(* IEC 61131-3 sources: JingjiangMoonbox/Application/Application/任务列表/OtherTask, 5 files *)

(* ---- KS_ArcFollow1UFlag_Deal.st ---- *)
(*@CES
Name=KS_ArcFollow1UFlag_Deal
Type=FunctionBlock
TypeGuid=6f9dac99-8de1-4efc-8465-68ac443b7d08
Guid=d7f43731-9672-42b8-a130-8c9a3b5ea44f
HasDeclaration=True
HasImplementation=True
*)
{DECLARATION}
FUNCTION KS_ArcFollow1UFlag_Deal : BOOL(*所有套色跟踪第一色标志处理@优化为了跟踪任意色@2024.02.22.102708*)
(*输出的标志可能决定了是否打开双波门*)
(*套色误差到达一定阈值时输出跟踪第一色标志-置位后就不再复位除非关闭使能
@用于解决在拉伸比较大的材料上后面色组找不到1色的问题。
@最大16个轴@c_byAxisNum_Max 确定*)
(*2024.02.22.085437 将检查第一个套色轴修改为检查跟踪的套色轴的下一个轴的误差*)
(*2025.1.9.145517 增加套色轴到达误差范围标志*)
VAR_INPUT
	i_xEn:BOOL;(*处理使能*)
	i_byArcNum_Max:BYTE;(*最大套色轴个数@最大16个*)
	i_byGrpAxisNum_Pu:BYTE;(*系中色组轴个数*)
	i_pabyGrpAxisList:POINTER TO BYTE;(*系的轴ID列表首地址*)
	i_byArcNum:BYTE;(*当前套色轴个数*)
	i_pabyArcAxisList:POINTER TO BYTE;(*套色的轴列表首地址@2024.02.22.084654*)
	i_pabyArcIdList:POINTER TO BYTE;(*套色的ID列表首地址*)
	i_byArcErr_Threshold:BYTE:=50;(*套色误差阈值@单位丝*)
	i_byContinuousCycleCnt:BYTE:=10;(*持续的圈数@持续这么多幅误差都在阈值以内就认为可以输出标志*)
	i_paxArcErrValid:POINTER TO ARRAY [1..c_byAxisNum_Max] OF BOOL;(*误差值有效了*)
	i_aiArcErr:ARRAY [1..c_byAxisNum_Max] OF INT;(*套色误差值(在让料头未到达的时候误差值写成最大值)@索引为色组号*)
	i_pabyCycleCnt:POINTER TO ARRAY [1..c_byAxisNum_Max] OF BYTE;(*满足条件后的圈数计数值@索引为色组号*)
	i_paxArcReachRangeFlag:POINTER TO ARRAY [1..c_byAxisNum_Max] OF BOOL;(*套色到达阈值标志@用于判断是否要输出跟踪第一色标志*)
	i_paxArcFollow1UFlag:POINTER TO ARRAY [1..c_byAxisNum_Max] OF BOOL;(*输出跟踪第一色标志@索引为色组号*)
	i_pabyFollowArcId:POINTER TO ARRAY [1..c_byAxisNum_Max] OF BYTE;(*2024.02.22.100117 跟踪的套色id@索引为轴id*)
	i_pxArcErrInRange:POINTER TO BOOL;(*套色误差在范围内@2025.1.9.145628+*)
END_VAR
VAR
	iN: INT;
	iM: INT;
	iAxisId: INT;
	iArcId: INT;
	byArcNum_Max: BYTE;
	byArcErr_Threshold: BYTE;(*丝单位*)
	byContinuousCycleCnt: BYTE;(*持续的幅数计数值*)

	byGrpAxisNum_Pu: BYTE;
	pabyGrpAxisList_Tmp:POINTER TO ARRAY [1..c_byAxisNum_Max] OF BYTE;(*系轴id列表*)
	abyGrpAxisList:ARRAY [1..c_byAxisNum_Max] OF BYTE;(*系轴id列表*)

	byArcNum: BYTE;
	pabyArcAxisList_Tmp:POINTER TO ARRAY [1..c_byAxisNum_Max] OF BYTE;(*套色轴id列表*)
	abyArcAxisList:ARRAY [1..c_byAxisNum_Max] OF BYTE;(*套色轴id列表*)
	pabyArcIdList_Tmp:POINTER TO ARRAY [1..c_byAxisNum_Max] OF BYTE;(*套色轴色序id列表*)
	abyArcIdList:ARRAY [1..c_byAxisNum_Max] OF BYTE;(*套色轴色序id列表*)
	axArcReachRangeFlag:ARRAY [1..c_byAxisNum_Max] OF BOOL;(*套色到达阈值标志*)
	axArcFollow1UFlag:ARRAY [1..c_byAxisNum_Max] OF BOOL;(*输出跟踪第一色标志@索引为色组号*)
	abyCycleCnt:ARRAY [1..c_byAxisNum_Max] OF BYTE;(*每个轴的循环计数*)
	aiArcErr:ARRAY [1..c_byAxisNum_Max] OF INT;(*套色误差*)
	axNeedRstAxisId: ARRAY [1..c_byAxisNum_Max] OF BOOL;(*需要复位参数的轴id|默认写true'*)
	axArcErrValid: ARRAY [1..c_byAxisNum_Max] OF BOOL;(*套色误差有效标志位*)
	xArvErrValid: BOOL;(*误差都有效了-可以检查标志*)
	xFollow1UEn: BOOL;(*跟踪第一色使能了*)

	abyFollowArcId:ARRAY [1..c_byAxisNum_Max] OF BYTE;(*2024.02.22.100 跟踪的套色id*)
	iFollowArcId:INT;
	iCheckArcIdSa:INT;(*开始检查的套色id*)
	iIndex: INT;
	iArcErrInRangeAxisCnt: INT;(*在范围的轴个数@2025.1.9.145758*)
END_VAR

VAR CONSTANT
	(*修改的时候谨慎点@外面输入的都是16个轴*)
	c_byAxisNum_Max:BYTE:=16;(*最大的轴个数@直接写死*)
END_VAR
{IMPLEMENTATION}
byArcNum_Max:=i_byArcNum_Max;
IF byArcNum_Max=0 OR
	byArcNum_Max>c_byAxisNum_Max THEN
	byArcNum_Max:=c_byAxisNum_Max;
END_IF

byArcNum:=i_byArcNum;
IF byArcNum>c_byAxisNum_Max THEN
	byArcNum:=c_byAxisNum_Max;
END_IF

byGrpAxisNum_Pu:=i_byGrpAxisNum_Pu;
IF byGrpAxisNum_Pu>c_byAxisNum_Max THEN
	byGrpAxisNum_Pu:=c_byAxisNum_Max;
END_IF

byArcErr_Threshold:=i_byArcErr_Threshold;
byContinuousCycleCnt:=i_byContinuousCycleCnt;

IF i_paxArcErrValid<>0 THEN
	axArcErrValid:=i_paxArcErrValid^;
END_IF
aiArcErr:=i_aiArcErr;

(*获取系轴列表信息*)
IF i_pabyGrpAxisList<>0 THEN
	pabyGrpAxisList_Tmp:=i_pabyGrpAxisList;
	abyGrpAxisList:=pabyGrpAxisList_Tmp^;
END_IF

(*获取套色轴列表信息*)
IF i_pabyArcAxisList<>0 THEN
	pabyArcAxisList_Tmp:=i_pabyArcAxisList;
	abyArcAxisList:=pabyArcAxisList_Tmp^;
END_IF

IF i_pabyArcIdList<>0 THEN
	pabyArcIdList_Tmp:=i_pabyArcIdList;
	abyArcIdList:=pabyArcIdList_Tmp^;
END_IF

IF i_pabyCycleCnt<>0 THEN
	abyCycleCnt:=i_pabyCycleCnt^;
END_IF
IF i_paxArcReachRangeFlag <>0 THEN
	axArcReachRangeFlag:=i_paxArcReachRangeFlag^;
END_IF
IF i_paxArcFollow1UFlag<>0 THEN
	axArcFollow1UFlag:=i_paxArcFollow1UFlag^;
END_IF

IF i_pabyFollowArcId<>0 THEN
	abyFollowArcId:=i_pabyFollowArcId^;
END_IF

(*只处理当前系的轴*)
FOR iN:=1 TO c_byAxisNum_Max BY 1 DO(*iN为系id索引*)
	iAxisId:=abyGrpAxisList[iN];
	IF iAxisId>0 AND iAxisId<c_byAxisNum_Max THEN
		axNeedRstAxisId[iAxisId]:=TRUE;
	ELSE;(*不在这个系的轴就不管了*)
	END_IF
END_FOR

iArcErrInRangeAxisCnt:=0;
FOR iN:=2 TO byArcNum BY 1 DO(*iN为索引@从第二个套色轴开始*)
	iAxisId:=abyArcAxisList[iN];(*套色的轴id*)
	iArcId:=abyArcIdList[iN];(*套色的色序id*)
	iFollowArcId:=abyFollowArcId[iN];(*跟踪的套色Id@2024.02.22.100304*)

	IF iAxisId>=2 AND iAxisId<=c_byAxisNum_Max AND(*轴号合法@从2号轴开始*)
		iArcId>=2 AND iArcId<=c_byAxisNum_Max THEN(*色序id合法*)
		xArvErrValid:=axArcErrValid[iAxisId];(*获取误差是否有效标志位*)
		axArcErrValid[iAxisId]:=FALSE;(*使用完了就复位*)
		(*检查各个色组是否到达阈值*)
		KS_ArcAxisReachRange(
			i_xEn (*i_xEn*),
			INT_TO_BYTE(iArcId)(*i_byArcId*),
			byArcErr_Threshold(*i_byArcErr_Threshold*),
			byContinuousCycleCnt(*i_byContinuousCycleCnt*),
			xArvErrValid(*i_xArcErrValid*),
			aiArcErr[iAxisId](*i_iArcErr*),
			ADR(abyCycleCnt[iAxisId])(*i_pbyCycleCnt*),
			ADR(axArcReachRangeFlag[iAxisId])(*i_xArcReachRangeFlag*));

		(*2025.1.9.145715+*)
		IF axArcReachRangeFlag[iAxisId] THEN
			iArcErrInRangeAxisCnt:=iArcErrInRangeAxisCnt+1;
		END_IF

		(*当前色已经到达阈值了@检查之前的套色轴是否到达。确定是否要输出跟踪第一色标志*)
		IF iFollowArcId<>0 THEN(*跟踪任意色@色序id*)
			IF iArcId>2 THEN(*色序超过3的才检查别的色*)
				IF axArcReachRangeFlag[iAxisId] THEN
					(*找到跟踪的套色id在套色id列表的索引值@2024.02.22.101030+*)
					iIndex:=iN;(*非法处理@未找到色序下面判断的循环就直接跳出*)
					FOR iM:=1 TO iN-1 BY 1 DO
						IF iFollowArcId = abyArcIdList[iM]THEN
							iIndex:=iM;
							EXIT;
						END_IF
					END_FOR

					(*如果找不到,会进入下面的else分支,但是iIndex=iN|所以也不会进入循环-也就是标志不会被置位*)
					iCheckArcIdSa:=2;
					IF iIndex<>In THEN(*找到了*)
						iIndex:=iIndex+1;(*从跟踪的下一个开始检查@索引值为开始检索的值*)
						iCheckArcIdSa:=abyArcIdList[iIndex];
					END_IF

					IF iCheckArcIdSa>=iArcId THEN(*检查的值和当前的色序一样@就直接输出标志*)
						axArcFollow1UFlag[iAxisId]:=TRUE;
					ELSE(*需要经过下面的检查输出*)
						(*修改为了跟踪色+1开始@2024.02.22.104458*)
						FOR iM:=iIndex TO iN-1  BY 1 DO(*从2色色序开始检查-自己在外围条件已经检查了@im也是色序*)
							IF axArcReachRangeFlag[abyArcAxisList[iM]] THEN(*到达阈值范围了*)
								IF iM=iN-1 THEN(*前一个也到达了则输出跟踪第一色标志*)
									axArcFollow1UFlag[iAxisId]:=TRUE;
								END_IF
							ELSE(*未到达则退出循环*)
								EXIT;
							END_IF
						END_FOR
					END_IF
				ELSE
					axArcFollow1UFlag[iAxisId]:=FALSE;
				END_IF
			ELSE
				axArcFollow1UFlag[iAxisId]:=axArcReachRangeFlag[iAxisId];(*只关心自己*)
			END_IF
		ELSE(*不跟踪任意色*)
			axArcFollow1UFlag[iAxisId]:=FALSE;
		END_IF
		(*处理未套色轴-复位标志@套色轴辅助变量已经在上面清除处理了*)
		axNeedRstAxisId[iAxisId]:=FALSE;
	ELSE;(*不做处理*)
	END_IF
END_FOR
(*检查所有轴是不是都在范围内@2025.1.9.145846*)
IF i_pxArcErrInRange<>0 THEN
	IF	(iArcErrInRangeAxisCnt+1) = byArcNum AND byArcNum>1 THEN
		i_pxArcErrInRange^:=TRUE;
	ELSE
		i_pxArcErrInRange^:=FALSE;
	END_IF
END_IF

(*没处理的轴数据清除*)
FOR iAxisId:=1 TO c_byAxisNum_Max BY 1 DO
	IF axNeedRstAxisId[iAxisId] THEN
		abyCycleCnt[iAxisId]:=0;
		axArcReachRangeFlag[iAxisId]:=FALSE;
		axArcFollow1UFlag[iAxisId]:=FALSE;
		axArcErrValid[iAxisId]:=FALSE;
	END_IF
END_FOR

IF i_pabyCycleCnt<>0 THEN
	i_pabyCycleCnt^:=abyCycleCnt;
END_IF
IF i_paxArcReachRangeFlag <>0 THEN
	i_paxArcReachRangeFlag^:=axArcReachRangeFlag;
END_IF
IF i_paxArcFollow1UFlag<>0 THEN
	i_paxArcFollow1UFlag^:=axArcFollow1UFlag;
END_IF

IF i_paxArcErrValid<>0 THEN
	i_paxArcErrValid^:=axArcErrValid;
END_IF

(* ---- KS_CalcGatePos_Follow.st ---- *)
(*@CES
Name=KS_CalcGatePos_Follow
Type=FunctionBlock
TypeGuid=6f9dac99-8de1-4efc-8465-68ac443b7d08
Guid=4fe415d3-d686-4f37-995a-ecb110eaba4a
HasDeclaration=True
HasImplementation=True
*)
{DECLARATION}
FUNCTION KS_CalcGatePos_Follow : INT(*计算跟踪某一个色方式计算该色的波门位置@单位是粗采样点数*)
(*-1 参数错误
-2 标记非法
-3 未隔色*)
(*2024.02.21.130156 输出第二波们的位置@出错则输出=0*)
(*2024.7.30.144846 计算方法有问题取巧未使用实际距离使用了波门宽度@波门宽度变化为非20后就会出错了
处理为根据实际距离计算*)
(*2024.7.31.075422 2色按照波门宽度偏移*)
VAR_INPUT
	i_byUnitId_Follow:BYTE;(*跟踪的色组id*)
	i_byUnitId_Cur:BYTE;(*当前的色组id*)
	i_iGateSa:INT;(*当前波门位置*)
	i_iGateWidthRondPt:INT;(*波门宽度的粗采样点数@使用改变量需要波门宽度为20mm*)
	i_iGatePoint_Max:INT;(*最大粗采样点数*)
	i_iMarkArrangeId:INT;(*标记类型*)

	i_rGirth:REAL;(*版辊周长@mm*)
END_VAR
VAR
	byDeltaId: BYTE;
	iGateSaEx: INT;
	iRtn: INT;
	iDeltaRondPt: INT;(*间隔的粗采样点数*)
END_VAR
{IMPLEMENTATION}
IF i_iGatePoint_Max=0 THEN
	i_iGatePoint_Max:=4000;
END_IF
IF i_byUnitId_Follow>0 AND
	i_byUnitId_Cur>=2 AND(*条件修改*)
	i_byUnitId_Follow<i_byUnitId_Cur AND
	i_iGateSa>=0 AND i_iGateSa<i_iGatePoint_Max THEN

	IF i_byUnitId_Cur>i_byUnitId_Follow THEN
		byDeltaId:=i_byUnitId_Cur-i_byUnitId_Follow;(*间隔*)
	ELSE
		byDeltaId:=0;
	END_IF

	IF byDeltaId<>0 THEN;
	ELSE(*不隔色*)
		iGateSaEx:= 0;
		iRtn:=-3;
		RETURN;
	END_IF

	IF i_rGirth<>0 THEN;
	ELSE
		i_rGirth:=500;
	END_IF
	IF i_byUnitId_Cur=2 THEN(*2色按照波门宽度偏移@2024.7.31.075310*)
		iDeltaRondPt:=i_iGateWidthRondPt;
	ELSE
		iDeltaRondPt:=REAL_TO_INT(BYTE_TO_REAL(byDeltaId)*20.0/i_rGirth*i_iGatePoint_Max)+1;(*按照间隔n*20mm计算|稍微离远点@主要是1 2色的波门*)
	END_IF

	IF i_iMarkArrangeId= MARK_ARRANGE_VFOR THEN(*顺序*)
		iGateSaEx:=i_iGateSa-(*byDeltaId*i_iGateWidthRondPt*)iDeltaRondPt;
		IF iGateSaEx<0 THEN
			iGateSaEx:= iGateSaEx+i_iGatePoint_Max;
		END_IF
	ELSIF i_iMarkArrangeId= MARK_ARRANGE_VREV THEN(*逆序*)
		iGateSaEx:=i_iGateSa+(*byDeltaId*i_iGateWidthRondPt*)iDeltaRondPt;
		IF iGateSaEx>i_iGatePoint_Max THEN
			iGateSaEx:= iGateSaEx-i_iGatePoint_Max;
		END_IF
	ELSE
		iGateSaEx:= 0;
		iRtn:=-2;
	END_IF
ELSE
	iGateSaEx:= 0;
	iRtn:=-1;
END_IF
(*
IF iRtn<0 THEN
	KS_CalcGatePos_Follow:=iRtn;
ELSE*)
	KS_CalcGatePos_Follow:=iGateSaEx;
(*END_IF*)

(* ---- KS_FB_GetLatchValue.st ---- *)
(*@CES
Name=KS_FB_GetLatchValue
Type=FunctionBlock
TypeGuid=6f9dac99-8de1-4efc-8465-68ac443b7d08
Guid=ed2f2b11-af18-4922-a052-26b8330b7fb0
HasDeclaration=True
HasImplementation=True
*)
{DECLARATION}
FUNCTION_BLOCK KS_FB_GetLatchValue
VAR_INPUT
	i_xEn : BOOL;
	i_iGrpUnitNum: INT;
	i_pstStSysParam: POINTER TO StSysParam;
	i_pastStLatch : POINTER TO ARRAY [1..MAX_UNIT_NUM] OF StLatch;
END_VAR
VAR_OUTPUT
END_VAR
VAR
	iN : INT;
	iM : INT;
	iRtn : INT;
	audiTempData : ARRAY [1..MAX_UNIT_NUM] OF UDINT;
END_VAR

{IMPLEMENTATION}

IF i_xEn THEN
	IF i_pstStSysParam <> 0 AND i_pastStLatch <> 0 THEN
		FOR iN := 1 TO i_iGrpUnitNum BY 1 DO
			iRtn := GTN_GetMailbox(
				core:= 1,
				station:= 0,
				byteAddress:= 16#C412, //锁存时间32位数据（低24位锁存时间，高8位di触发次数），单位us,:低16位网络地址0xc412,高16位网络地址0xc414
				pData:= ADR(audiTempData[iN]),
				wordCount:= 2,
				dataMode:= 1,
				desId:=iN,
				typeVar:= 1);

			i_pastStLatch^[iN].iTriggerCnt := UDINT_TO_INT(SHR(audiTempData[iN],24));
			i_pastStLatch^[iN].udiTriggerTimeErr := SHR(SHL(audiTempData[iN],16#8),16#8);

			iRtn := GTN_GetMailbox(
				core:= 1,
				station:= 0,
				byteAddress:= 16#C454, //锁存编码器32位数据，一个版周最大脉冲值131072，低16位网络地址0xc454，高16位网络地址0xc456
				pData:= ADR(i_pastStLatch^[iN].udiTriggerEncErr),
				wordCount:= 2,
				dataMode:= 1,
				desId:=iN,
				typeVar:= 1);
		END_FOR
	END_IF
ELSE
	;
END_IF

(* ---- PRG_MODBUS_TCP.st ---- *)
(*@CES
Name=PRG_MODBUS_TCP
Type=FunctionBlock
TypeGuid=6f9dac99-8de1-4efc-8465-68ac443b7d08
Guid=8040f7c3-2c5c-428c-829e-f8dbe8b2490b
HasDeclaration=True
HasImplementation=True
*)
{DECLARATION}
PROGRAM PRG_MODBUS_TCP
VAR
	axCoils: ARRAY [1..2] OF BYTE;(*线圈*)
	axDiscreteInput: ARRAY [1..2] OF BYTE;(*离散线圈*)
	awInputReg: ARRAY [1..2] OF WORD;(*输入寄存器*)
	awHoldingReg: ARRAY [1..1000] OF WORD;(*保持寄存器区*)
	wPort_VisionUI: WORD := 502;(*视觉访问的端口号*)
	udiXOFST_VisionUIGave: UDINT := 0;(*4字节*)
	uiXOFST_UpdateFlag: UINT := 0;(*X坐标值被更新标志*)
	//fbModbus_TCP_Slave: Modbus_TCP_Slave;(*ModBus TCP从站功能*)

	dwGirth_Temp:DWORD;
	wGirth_Temp_L:WORD;
	wGirth_Temp_H:WORD;
		(*地址约定
		40116: X坐标测量功能的使能,=1表示可以采集,其余值(推荐0)均为不可以.科赛程序控制;固德只读;
		40871: 测量X坐标的偏差(数据低位);固德写给科赛;
		40872: 测量X坐标的偏差(数据高位);固德写给科赛;
		40873: 写1表示40871和40872被更新了;科赛读取数据后写0即可
		40007: 版周长低位
		40008: 版周长高位
		*)
END_VAR

{IMPLEMENTATION}
awHoldingReg[116]:= BOOL_TO_WORD(g_xSendResToOnline);(*使能标志*)
//2026.04.11.184336 增加版周长通讯
dwGirth_Temp:=REAL_TO_DWORD(g_stStSysParam.astStGrpParam_Save[1].rGirth_PrnRoller*1000);
wGirth_Temp_L:=DWORD_TO_WORD(dwGirth_Temp);
wGirth_Temp_H:=DWORD_TO_WORD(SHR(dwGirth_Temp,16));
awHoldingReg[7]:=wGirth_Temp_L;
awHoldingReg[8]:=wGirth_Temp_H;
(*
fbModbus_TCP_Slave(
	pCoils:= ADR(axCoils),
	pDiscreteInput:= ADR(axDiscreteInput),
	pInputReg:= ADR(awInputReg),
	pHoldingReg:= ADR(awHoldingReg),
	CMax:= 16,
	DIMax:= 16,
	IRMax:= 2,
	HRMax:= 1000,
	Enable:= TRUE,
	port:= wPort_VisionUI,
	Enable_WatchDog:= FALSE,
	tWatchDogTime:= ,
	ClientStatus=> ,
	wErrorId=> ,
	bError=> );
	*)
uiXOFST_UpdateFlag:= awHoldingReg[873];
IF uiXOFST_UpdateFlag=1 THEN
	g_stStSysParam.astStRSV_GrpParam_UnSave[1].xBasePosDoneByOnline:=TRUE;
	awHoldingReg[873]:=0;
	udiXOFST_VisionUIGave:= SHL(WORD_TO_UDINT(awHoldingReg[871]),16) OR WORD_TO_UDINT(awHoldingReg[872]);
	g_stStSysParam.astStRSV_GrpParam_UnSave[1].rFiberMoveBasePosByOnline:=UDINT_TO_REAL(udiXOFST_VisionUIGave)*0.001165+103.8341;

END_IF

(* ---- PRG_OTHER.st ---- *)
(*@CES
Name=PRG_OTHER
Type=FunctionBlock
TypeGuid=6f9dac99-8de1-4efc-8465-68ac443b7d08
Guid=e1db0700-f403-46d4-96bb-1521e027fd26
HasDeclaration=True
HasImplementation=True
*)
{DECLARATION}
PROGRAM PRG_OTHER
VAR
	iRtn : INT;
	iGrp : INT;
	iK : INT;
	iN : INT;
	iAxisId:INT;
	byColorId:BYTE;
	abyColorId_Bak:ARRAY [1..MAX_UNIT_NUM] OF BYTE;(*色序id备份值@2024.02.27.151112*)
	axInitValue_ClorId_Bak:ARRAY [1..2] OF BOOL;(*初始化色组id备份值@2024.02.27.151956*)
	abyGrpAxisNum_Pu: ARRAY [1..2] OF BYTE;

	pstStUnitParam_Save : POINTER TO StUnitParam_Save;
	pstStUnitParam_UnSave : POINTER TO StUnitParam_UnSave;

	pstStGrpParam_Save : POINTER TO StGrpParam_Save;
	pstStGrpParam_UnSave : POINTER TO StGrpParam_UnSave;

	abyNeedFollow_1U: ARRAY [1..2] OF BYTE;(*.0 纵向打开双波门
						    .1 横向打开双波门*)
	(*按系分*)
	axInitValue_FlagFollow_Bak: ARRAY [1..2] OF BOOL;(*初始化跟踪方式备份值@2024.02.27.151956*)
	abyLastNeedFollow_1U: ARRAY [1..2] OF BYTE;(*.0 纵向打开双波门
											 .1 横向打开双波门*)
	axInitValue_HorOpen_Bak: ARRAY [1..2] OF BOOL;(*横向打开备份值初始化@2024.02.27.154613*)
	axHorOpen_Bak:ARRAY [1..MAX_UNIT_NUM] OF BOOL;(*横向开关备份变量@2024.02.27.154642*)
	pbyTmp: POINTER TO BYTE;

	axAtLeastOneUnitOpenHor: ARRAY [1..2] OF BOOL;(*至少一色打开横向了*)

	(*2024.02.21.125231 优化跟踪第一色实现为任意色*)
	byFollowArcId: BYTE;

	(*2023.12.05.135403 跟踪第一色标志处理需要变量*)
	aiArcErr: ARRAY [1..16] OF INT;
	abyCycleCnt: ARRAY [1..16] OF BYTE;
	axArcReachRangeFlag: ARRAY [1..16] OF BOOL;
	axArcFollow1UFlag_WaitFilmLenth:  ARRAY [1..16] OF BOOL;(*等料长置位的跟一色标志*)
	axArcFollow1UFlag_ErrReachRange:  ARRAY [1..16] OF BOOL;(*误差到达一定范围以后才输出的置位标志*)

//	fbGT_GetSystemInfo : GT_GetSystemInfo;
	udiRemain_M : UDINT;
	iCount_1_Second : INT;
	xChangeSignal : BOOL;

	fbKS_FB_GetLatchValue : KS_FB_GetLatchValue;

	//2025.11.16.090955 | 获取CPU以及内存信息
	test_info:SystemInfo;
    plc_info:POINTER TO TSysInfo;

	uliRemain_M : ULINT;
	sPath : STRING;
	iCount_GetPlcInfo : INT;
//	iCount_GetPlcInfo : INT;
	iCount_DeleteDir : INT;
	byArcIntensity_Pre: BYTE;
	xChange_ArcIntensity: BOOL;
END_VAR

{IMPLEMENTATION}
IF g_iRunStepId=RUNSTEP_NormalWork THEN
	;
ELSE
	RETURN;
END_IF
g_stStSysParam.stStSysParam_Save.byTypeFollow1UEn:=1;

FOR iN:=1 TO MAX_UNIT_NUM BY 1 DO
	IF g_stStSysParam.astStUnitParam_Save[iN].rGirth_Sam <> 0 THEN
		g_stStSysParam.astStUnitParam_Save[iN].iGateWidthRoundPoints:=
				REAL_TO_INT(20.0/g_stStSysParam.astStUnitParam_Save[iN].rGirth_Sam*4000.0);
	ELSE
		g_stStSysParam.astStUnitParam_Save[iN].rGirth_Sam := g_stStSysParam.astStUnitParam_Save[iN].rGirth_PrnRoller;
	END_IF
END_FOR

(*2023.09.10.122156 优化*)
(*2024.02.21.125747 优化为跟踪任意色而不是单单跟踪第一色@变量名有点混淆.eg xFlag_Follow_1U_V 现在的意义是跟踪任意色*)
FOR iGrp:=1 TO 2 BY 1 DO
	pstStGrpParam_Save:=ADR(g_stStSysParam.astStGrpParam_Save[iGrp]);
	pstStGrpParam_UnSave:=ADR(g_stStSysParam.astStGrpParam_UnSave[iGrp]);
	abyGrpAxisNum_Pu[iGrp]:=pstStGrpParam_UnSave^.byGrpAxisNum_Pu;(*2023.09.21.135454 缺失了一段代码*)
	(*2023.11.27.102831 xFlag_Follow_1U_V的内存区域和之前使用的有点冲突，
	会引起xFlag_Follow_1U_V高位字节非零在这里强制清零处理只保留最低位*)
	pbyTmp:=ADR(pstStGrpParam_Save^.xFlag_Follow_1U_V);
	IF pbyTmp^>1 THEN(*非0 非1*)
		pbyTmp^:=pbyTmp^ AND 16#01;(*保留最低位*)
	END_IF
	(*检查至少一色横向打开了*)
	axAtLeastOneUnitOpenHor[iGrp]:=FALSE;
	FOR iK:=1 TO abyGrpAxisNum_Pu[iGrp] BY 1 DO
		iAxisId:=pstStGrpParam_UnSave^.abyGrpAxisList[iK];
		IF iAxisId>0 AND iAxisId<=MAX_UNIT_NUM THEN
			pstStUnitParam_Save:=ADR(g_stStSysParam.astStUnitParam_Save[iAxisId]);(*取轴参数*)
			pstStUnitParam_UnSave:=ADR(g_stStSysParam.astStUnitParam_UnSave[iAxisId]);(*取轴参数*)
			byColorId:=pstStUnitParam_UnSave^.byColorIdCurrent;(*取色序id*)
			IF byColorId>1 THEN(*色序大于1@只检测套印轴*)
				IF pstStUnitParam_Save^.dwFlag_Ctl.0 THEN(*至少打开了一个颜色的横向*)
					axAtLeastOneUnitOpenHor[iGrp]:=TRUE;
					EXIT;
				END_IF
			END_IF
		END_IF
	END_FOR

	abyNeedFollow_1U[iGrp]:=0;
	abyNeedFollow_1U[iGrp].0:=pstStGrpParam_Save^.xFlag_Follow_1U_V;(*打开纵向跟1色开关*)
	abyNeedFollow_1U[iGrp].1:=pstStGrpParam_Save^.xFlag_Follow_1U_H (*AND xAtLeastOneUnitOpenHor*);(*至少一色横向打开并且横向跟1色*)

	IF NOT axInitValue_FlagFollow_Bak[iGrp] THEN
		abyLastNeedFollow_1U[iGrp]:= abyNeedFollow_1U[iGrp];
		axInitValue_FlagFollow_Bak[iGrp]:=TRUE;

	END_IF

	FOR iK:=1 TO abyGrpAxisNum_Pu[iGrp] BY 1 DO
		iAxisId:=pstStGrpParam_UnSave^.abyGrpAxisList[iK];
		IF iAxisId>0 AND iAxisId<=MAX_UNIT_NUM THEN
			pstStUnitParam_Save:=ADR(g_stStSysParam.astStUnitParam_Save[iAxisId]);(*取轴参数*)
			pstStUnitParam_UnSave:=ADR(g_stStSysParam.astStUnitParam_UnSave[iAxisId]);(*取轴参数*)
			byColorId:=pstStUnitParam_UnSave^.byColorIdCurrent;(*取色序id*)

			(*跟踪的色序id进行处理@2024.02.27.152243*)
			IF NOT axInitValue_ClorId_Bak[iGrp] THEN
				abyColorId_Bak[iAxisId]:=byColorId;
				IF iK=abyGrpAxisNum_Pu[iGrp] THEN
					axInitValue_ClorId_Bak[iGrp]:=TRUE;(*循环完成了*)
				END_IF
			END_IF

			IF NOT axInitValue_HorOpen_Bak[iGrp] THEN
				axHorOpen_Bak[iAxisId]:=pstStUnitParam_Save^.dwFlag_Ctl.0;
				IF iK= abyGrpAxisNum_Pu[iGrp] THEN
					axInitValue_HorOpen_Bak[iGrp]:=TRUE;(*循环完成了*)
				END_IF
			END_IF

			(*横向跟任意色打开了|跟踪色未分配则写成1*)
			IF (abyLastNeedFollow_1U[iGrp] <> abyNeedFollow_1U[iGrp] AND abyNeedFollow_1U[iGrp].1) OR
				(*色序id从0变未非0,并且横向跟任意色打开,初始化跟踪色序*)
				(abyColorId_Bak[iAxisId]<>byColorId AND abyColorId_Bak[iAxisId]=0 AND abyNeedFollow_1U[iGrp].1) OR
				(*横向打开的时候并且横向跟任意色打开,初始化跟踪色序*)
				(NOT axHorOpen_Bak[iAxisId] AND pstStUnitParam_Save^.dwFlag_Ctl.0 AND abyNeedFollow_1U[iGrp].1) THEN
				IF pstStUnitParam_Save^.byFollowColorId=0 AND pstStUnitParam_Save^.dwFlag_Ctl.0 THEN(*=0 以及横向打开的轴强制写1*)
					pstStUnitParam_Save^.byFollowColorId:=1;
				END_IF
			END_IF

			(*2024.02.21.130709 关闭跟踪任意一色@强制将色组修改为跟踪前一色-双眼*)
			IF (abyLastNeedFollow_1U[iGrp] <> abyNeedFollow_1U[iGrp] AND abyNeedFollow_1U[iGrp]=0) OR
				byColorId<=1 OR(*色序id*)
				(*在纵向跟任意色未打开,横向跟踪任意色打开而横向开关打开时-强制followid=0*)
				(NOT abyNeedFollow_1U[iGrp].0 AND abyNeedFollow_1U[iGrp].1 AND NOT pstStUnitParam_Save^.dwFlag_Ctl.0) THEN
				pstStUnitParam_Save^.byFollowColorId:=0;
			END_IF

			(*检查当前色序id是否非法@超过当前色序则写0*)
			IF pstStUnitParam_Save^.byFollowColorId >= byColorId THEN
				pstStUnitParam_Save^.byFollowColorId:=0;(*强制写0*)
			END_IF

			IF g_stStSysParam.stStSysParam_Save.xArcFollowAnyAxis THEN;(*跟踪任意色|则由上面逻辑调整跟踪轴id*)
			ELSE(*只能跟踪第一色*)
				pstStUnitParam_Save^.byFollowColorId:=1;(*强制跟踪第一色@如果要跟踪任意色-屏蔽这行代码@2024.02.27.160908*)
			END_IF
			(*--END*)

			byFollowArcId:=pstStUnitParam_Save^.byFollowColorId;(*取跟踪的色id*)

			IF abyNeedFollow_1U[iGrp]<>0 THEN(*需要跟踪第一色*)
				IF byColorId>1 THEN(*色序大于1*)
					(*位状态处理@2023.09.10.214936*)
					IF abyNeedFollow_1U[iGrp].0 THEN(*纵向跟踪第一色*)
						IF byFollowArcId<>0 THEN(*跟踪的色序id非0则打开*)
							pstStUnitParam_Save^.dwFlag_Sts.8:= TRUE;
						ELSE(*跟踪色序为0的时候关闭*)
							pstStUnitParam_Save^.dwFlag_Sts.8:= FALSE;
						END_IF
					ELSE
						IF abyLastNeedFollow_1U[iGrp].0 THEN(*之前跟踪第一色按钮打开过*)
							pstStUnitParam_Save^.dwFlag_Sts.8:= FALSE;
						END_IF
					END_IF
					IF abyNeedFollow_1U[iGrp].1 THEN(*横向跟踪第一色*)
						IF byFollowArcId<>0 THEN(*跟踪的色序id非0则打开*)
							pstStUnitParam_Save^.dwFlag_Sts.9:= pstStUnitParam_Save^.dwFlag_Ctl.0;(*打开横向才置位*)
						ELSE(*跟踪色序为0的时候关闭*)
							pstStUnitParam_Save^.dwFlag_Sts.9:= FALSE;
						END_IF
					ELSE
						IF abyLastNeedFollow_1U[iGrp].1 THEN(*之前跟踪第一色按钮打开过*)
							pstStUnitParam_Save^.dwFlag_Sts.9:= FALSE;
						END_IF
					END_IF

					(*计算第二个波门位置@纵横向有一个打开跟踪第一色，第二波门自动计算*)
					pstStUnitParam_Save^.iGateSaEx:=
						KS_CalcGatePos_Follow(
							byFollowArcId(*i_byUnitId_Follow*),
							byColorId(*i_byUnitId_Cur*),
							pstStUnitParam_Save^.iGateSa(*i_iGateSa*),
							pstStUnitParam_Save^.iGateWidthRoundPoints(*i_iGateWidthRondPt*)+1,(*不要挨得太近+1个点*)
							4000(*i_iGatePoint_Max*),
							(*2024.03.06.171730 将整机的标记形式修改为了轴的标记形式*)
							pstStUnitParam_Save^.iMarkArrangeMode,(*pstStGrpParam^.iMarkArrangeId*)(*i_iMarkArrangeId*)
							pstStUnitParam_Save^.rGirth_PrnRoller(*i_rGirth*));
				ELSE(*色序为1就取消吧*)
					pstStUnitParam_Save^.dwFlag_Sts.8:= FALSE;
					pstStUnitParam_Save^.dwFlag_Sts.9:= FALSE;
					pstStUnitParam_Save^.iGateSaEx:=0;
				END_IF
			ELSE(*不需要跟踪第一色|根据界面选择控制*)
				IF abyLastNeedFollow_1U[iGrp].0 THEN(*之前跟踪第一色按钮打开过*)
					pstStUnitParam_Save^.dwFlag_Sts.8:= FALSE;
				END_IF
				IF abyLastNeedFollow_1U[iGrp].1 THEN(*之前跟踪第一色按钮打开过*)
					pstStUnitParam_Save^.dwFlag_Sts.9:= FALSE;
				END_IF
			END_IF

			(*纵横向都没有打开全跟踪第一色开关，第二波门手动指定*)
			IF pstStUnitParam_Save^.dwFlag_Sts.8 OR(*纵向跟踪任意一色*)
				pstStUnitParam_Save^.dwFlag_Sts.9 THEN(*横向跟踪任意一色*)
				(*打开双波门开关*)
				IF pstStUnitParam_Save^.iMarkArrangeMode=MARK_ARRANGE_OMK OR(*单标记*)
					pstStUnitParam_Save^.iMarkArrangeMode=MARK_ARRANGE_HFOR OR(*横顺*)
					pstStUnitParam_Save^.iMarkArrangeMode=MARK_ARRANGE_HREV THEN(*横逆*)
					pstStUnitParam_Save^.dwFlag_Ctl.6:=FALSE;(*不能打开双波门*)
				ELSE
					pstStUnitParam_Save^.dwFlag_Ctl.6:=TRUE;(*双波门标志有效*)
				END_IF
			ELSE
				pstStUnitParam_Save^.dwFlag_Ctl.6:= FALSE;(*双波门取消使能|强制关闭吧，反正界面打开计算误差哪里也没处理*)
			END_IF

			(*2023.09.14.103752 处理纵向使用哪一个误差进行计算调整量@处理开机时候pe裁切拉伸引起的找不到第一色问题
			在开机时候先使用跟踪前一色-随后切换未跟踪第一色*)

(*2023.12.05.135650  重新实现*)
(*
			IF pstStAxisParam^.wStatusRef.8 THEN(*跟第一色打开了*)
				IF pstStAxisParam^.xWaitFilmLenth_Follow1U THEN(*第一色没来的时候|先用跟踪前一色@xWaitFilmLenth_Follow1U=true正在等一色*)
					pstStAxisParam^.wStatusRef.12:=FALSE;(*使用跟踪前一色的误差计算调整量*)
				ELSE(*xWaitFilmLenth_Follow1U等完后会变成false*)
					pstStAxisParam^.wStatusRef.12:=TRUE;(*使用跟踪第一色的误差计算调整量*)
				END_IF
			ELSE
				pstStAxisParam^.wStatusRef.12:=FALSE;(*使用跟踪前一色的误差计算调整量*)
			END_IF
*)
			(*2023.12.05.135707 使能位更换为了局部变量*)
			IF iAxisId>=1 AND iAxisId<=16 THEN(*只处理前16个轴*)
				IF pstStUnitParam_Save^.dwFlag_Sts.8 THEN(*跟第一色打开了*)
					IF pstStUnitParam_Save^.xWaitFilmLenth_Follow1U THEN(*第一色没来的时候|先用跟踪前一色@xWaitFilmLenth_Follow1U=true正在等一色*)
						axArcFollow1UFlag_WaitFilmLenth[iAxisId]:=FALSE;(*使用跟踪前一色的误差计算调整量*)
					ELSE(*xWaitFilmLenth_Follow1U等完后会变成false*)
						axArcFollow1UFlag_WaitFilmLenth[iAxisId]:=TRUE;(*使用跟踪第一色的误差计算调整量*)
					END_IF
				ELSE
					axArcFollow1UFlag_WaitFilmLenth[iAxisId]:=FALSE;(*使用跟踪前一色的误差计算调整量*)
				END_IF
			END_IF
		END_IF
		abyColorId_Bak[iAxisId]:=byColorId;(*2024.02.27.151208 +*)
		axHorOpen_Bak[iAxisId]:=pstStUnitParam_Save^.dwFlag_Ctl.0;
	END_FOR
	abyLastNeedFollow_1U[iGrp]:=abyNeedFollow_1U[iGrp];(*打开过跟一色*)

	(*按照系循环*)
	(*2023.12.05.135016 跟踪第一色标志处理@前面色组误差到达一定阈值后输出标志*)
	SysMemCpy(ADR(aiArcErr),ADR(g_aiArcErr_V),SIZEOF(aiArcErr));(*误差拷贝*)
	KS_ArcFollow1UFlag_Deal(
		pstStGrpParam_UnSave^.xFlag_Print AND(*印刷状态|速度大于10*)
		pstStGrpParam_UnSave^.rVel_Film>=10 (*AND(*印刷状态|速度大于10*)
		pstStGrpParam^.xFlag_Follow_1U_V*)(*i_xEn*),(*打开了跟踪第一色*)(*2025.1.9.150129 有效了就使能*)
		16(*i_byArcNum_Max*),
		pstStGrpParam_UnSave^.byGrpAxisNum_Pu(*i_byGrpAxisNum_Pu*),
		ADR(pstStGrpParam_UnSave^.abyGrpAxisList)(*i_pabyGrpAxisList*),
		pstStGrpParam_UnSave^.byGrpArcAxisNum(*i_byArcNum*),
		ADR(pstStGrpParam_UnSave^.abyGrpArcAxisList)(*i_pabyArcAxisList*),
		ADR(pstStGrpParam_UnSave^.abyGrpArcIdList)(*i_pabyArcIdList*),
		(*2025.1.10.122923 判断误差稳定的阈值修改到1mm*)
		100(*i_byArcErr_Threshold*),
		10(*i_byContinuousCycleCnt*),
		ADR(g_axArcErrValid)(*i_paxArcErrValid*),(*等料长完成后一圈会置位一次@只处理了前16个id索引*)
		aiArcErr(*i_aiArcErr*),
		ADR(abyCycleCnt)(*i_pabyCycleCnt*),
		ADR(axArcReachRangeFlag)(*i_paxArcReachRangeFlag*),
		ADR(axArcFollow1UFlag_ErrReachRange)(*i_paxArcFollow1UFlag*),
		ADR(pstStGrpParam_UnSave^.abyGrpFollowArcIdList)(*i_pabyFollowArcId*),
		ADR(pstStGrpParam_UnSave^.xArcErrInRange)(*i_pxArcErrInRange*));

	FOR iK:=1 TO abyGrpAxisNum_Pu[iGrp] BY 1 DO
		iAxisId:=pstStGrpParam_UnSave^.abyGrpAxisList[iK];
		IF iAxisId>0 AND iAxisId<=16 THEN(*只处理前16个轴*)
			pstStUnitParam_Save:=ADR(g_stStSysParam.astStUnitParam_Save[iAxisId]);(*取轴参数*)
			pstStUnitParam_UnSave:=ADR(g_stStSysParam.astStUnitParam_UnSave[iAxisId]);(*取轴参数*)
			(*安全起见 and pstStAxisParam^.wStatusRef.8*)
			CASE g_stStSysParam.stStSysParam_Save.byTypeFollow1UEn OF
				1:(*等料长结束了就切换*)
					pstStUnitParam_Save^.dwFlag_Sts.12:=axArcFollow1UFlag_WaitFilmLenth[iAxisId] AND pstStUnitParam_Save^.dwFlag_Sts.8;
				2:(*直接使能@2024.03.21.102817*)
					pstStUnitParam_Save^.dwFlag_Sts.12:=pstStUnitParam_Save^.dwFlag_Sts.8;
			ELSE(*等料长结束后-等待前色误差进入阈值范围内切换*)
					(*2024.9.3.092214 优化为了1色料长到了强制转换*)
(*					pstStAxisParam^.wStatusRef.12:=pstStAxisParam^.wStatusRef.8 AND
							(axArcFollow1UFlag_ErrReachRange[iAxisId] OR axArcFollow1UFlag_WaitFilmLenth[iAxisId]);*)
					pstStUnitParam_Save^.dwFlag_Sts.12:=pstStUnitParam_Save^.dwFlag_Sts.8 AND
							(axArcFollow1UFlag_ErrReachRange[iAxisId]);
			END_CASE

			IF (pstStGrpParam_UnSave^.xFlag_Ink AND pstStGrpParam_UnSave^.xEnaTestARC_Ink) THEN(*空转单眼调试*)
				pstStUnitParam_Save^.dwFlag_Sts.12:=pstStUnitParam_Save^.dwFlag_Sts.8;(*如果选择跟踪第一色，就直接赋值*)
			END_IF

			(*2024.01.02.113642 同步*)
			(*2023.12.25.212750+持续一定时间后结束*)
			IF pstStGrpParam_UnSave^.xFlag_Follow_1U_V_UwCut OR
				pstStGrpParam_UnSave^.xFlagFollow1U_AccDecing THEN(*2024.04.14.114538+*)
				pstStUnitParam_Save^.dwFlag_Sts.12:=TRUE;(*接料时候跟踪第一色计算误差*)
				IF pstStUnitParam_Save^.iMarkArrangeMode=MARK_ARRANGE_OMK OR(*单标记*)
					pstStUnitParam_Save^.iMarkArrangeMode=MARK_ARRANGE_HFOR OR(*横顺*)
					pstStUnitParam_Save^.iMarkArrangeMode=MARK_ARRANGE_HREV THEN(*横逆*);
				ELSE;
					pstStUnitParam_Save^.dwFlag_Ctl.6:=TRUE;(*打开双波门*)
				END_IF
			END_IF
		END_IF
	END_FOR

	(*2024.8.30.102618增加全控双眼/单眼跟1色开关*)
	FOR iK:=1 TO abyGrpAxisNum_Pu[iGrp] BY 1 DO
		iAxisId:=pstStGrpParam_UnSave^.abyGrpAxisList[iK];
		IF iAxisId>0 AND iAxisId<=16 THEN(*只处理前16个轴*)
			pstStUnitParam_Save:=ADR(g_stStSysParam.astStUnitParam_Save[iAxisId]);(*取轴参数*)
			pstStUnitParam_UnSave:=ADR(g_stStSysParam.astStUnitParam_UnSave[iAxisId]);(*取轴参数*)
			pstStUnitParam_Save^.dwFlag_Sts.14:= g_stStSysParam.stStSysParam_Save.xFlag_Follow_1U_Double_V;
			pstStUnitParam_Save^.dwFlag_Sts.15:= g_stStSysParam.stStSysParam_Save.xFlag_Follow_1U_Double_H;
		END_IF
	END_FOR
END_FOR

//2025.11.6.140503保存系统配置按钮|niuj
IF g_xBtn_UpdateSysCfg THEN
	g_xBtn_UpdateSysCfg:= FALSE;
	g_xInit_TrapPoint:= FALSE;
	IF g_stStSysParam.astStGrpParam_UnSave[1].xFlag_Stop OR
		g_stStSysParam.astStGrpParam_UnSave[2].xFlag_Stop OR
		g_stStSysParam.astStGrpParam_UnSave[1].xFlag_EStop OR
		g_stStSysParam.astStGrpParam_UnSave[2].xFlag_EStop THEN

// 		SysMemCpy(
// 				ADR(g_stStSysParam.stStSysParam_UnSave.stStSysCfgStruct),
// 				ADR(g_stStSysCfgStruct),
// 				SIZEOF(g_stStSysCfgStruct));
		g_iRunStepId:= RUNSTEP_UpdateSysCfg;
		g_xInit_StationList := FALSE;
	END_IF

END_IF

//2025.11.16.090955 | 获取CPU以及内存信息
iCount_GetPlcInfo := iCount_GetPlcInfo + 1;
IF iCount_GetPlcInfo > 9 THEN
	iCount_GetPlcInfo := 0;
	test_info(PLC_SYS_INFO => plc_info);
	uliRemain_M := plc_info^.space_info[5].remain/1024/1024;
	FOR iN := 0 TO 3 BY 1 DO
		g_abyCpu_Load[iN] := REAL_TO_BYTE(plc_info^.CPU_Load[iN]);
	END_FOR

	IF uliRemain_M < 1000 THEN
		iCount_DeleteDir := iCount_DeleteDir + 1;
		IF iCount_DeleteDir > 19 THEN
			iCount_DeleteDir := 0;
			sPath :=  '/data/kesai/data';
			GTN_KSDirDelete(file:= ADR(sPath));
		END_IF
	ELSE
		iCount_DeleteDir := 0;
	END_IF
END_IF

iCount_1_Second := iCount_1_Second+1;
IF iCount_1_Second >= 10 THEN
	IF NOT xChangeSignal THEN
		xChangeSignal := TRUE;
		g_sHandConnectedSignal := '#';
	ELSE
		xChangeSignal := FALSE;
		g_sHandConnectedSignal := ' ';
	END_IF
END_IF

//2025.12.26.112513 | 获取锁存的内容，临时先放在这个任务当中，因为目前的MailBox获取方法耗时比较长
fbKS_FB_GetLatchValue(
	i_xEn:= FALSE,
	i_iGrpUnitNum:= g_stStSysParam.astStGrpParam_UnSave[1].byGrpAxisNum_Pu,
	i_pstStSysParam:= ADR(g_stStSysParam),
	i_pastStLatch:= ADR(g_astStLatch)
	);

(*2026.4.25.145102处理界面调整强度切换*)
IF g_stStSysParam.stStSysParam_Save.byArcIntensity_W= 0 THEN
	g_stStSysParam.stStSysParam_Save.byArcIntensity_W:= 25;
END_IF

IF g_stStSysParam.stStSysParam_Save.byArcIntensity_M= 0 THEN
	g_stStSysParam.stStSysParam_Save.byArcIntensity_M:= 20;
END_IF

IF g_stStSysParam.stStSysParam_Save.byArcIntensity_S= 0 THEN
	g_stStSysParam.stStSysParam_Save.byArcIntensity_S:= 15;
END_IF

//新增套色强度切换逻辑2026.4.25.150042||
IF g_stStSysParam.stStSysParam_Save.byArcIntensity<>byArcIntensity_Pre THEN
	xChange_ArcIntensity:= TRUE;
END_IF
byArcIntensity_Pre:= g_stStSysParam.stStSysParam_Save.byArcIntensity;
IF xChange_ArcIntensity THEN
	xChange_ArcIntensity:= FALSE;
	FOR iN:=1 TO MAX_UNIT_NUM BY 1 DO
		IF g_stStSysParam.stStSysParam_Save.byArcIntensity=0 THEN
			g_stStSysParam.astStUnitParam_Save[iN].rMargin_Mag_Arc:= g_stStSysParam.stStSysParam_Save.byArcIntensity_W;
			g_stStSysParam.astStUnitParam_Save[iN].stStArc_Mol_Param.rMargin_Mag_Arc:= g_stStSysParam.stStSysParam_Save.byArcIntensity_W;
		ELSIF g_stStSysParam.stStSysParam_Save.byArcIntensity=1 THEN
			g_stStSysParam.astStUnitParam_Save[iN].rMargin_Mag_Arc:= g_stStSysParam.stStSysParam_Save.byArcIntensity_M;
			g_stStSysParam.astStUnitParam_Save[iN].stStArc_Mol_Param.rMargin_Mag_Arc:= g_stStSysParam.stStSysParam_Save.byArcIntensity_M;
		ELSIF g_stStSysParam.stStSysParam_Save.byArcIntensity=2 THEN
			g_stStSysParam.astStUnitParam_Save[iN].rMargin_Mag_Arc:= g_stStSysParam.stStSysParam_Save.byArcIntensity_S;
			g_stStSysParam.astStUnitParam_Save[iN].stStArc_Mol_Param.rMargin_Mag_Arc:= g_stStSysParam.stStSysParam_Save.byArcIntensity_S;
		ELSE
			g_stStSysParam.astStUnitParam_Save[iN].rMargin_Mag_Arc:= g_stStSysParam.stStSysParam_Save.byArcIntensity_M;
			g_stStSysParam.astStUnitParam_Save[iN].stStArc_Mol_Param.rMargin_Mag_Arc:= g_stStSysParam.stStSysParam_Save.byArcIntensity_M;

		END_IF
	END_FOR
END_IF
